// TIA Portal V20 export
// export: Created 2026-10-19T18:01:35.4601049Z, ExportSetting None, DisplayName Totally Integrated Automation Portal, DisplayVersion V20 Update 6, DisplayName TIA Portal Openness, DisplayVersion V20 Update 6, DisplayName TIA Portal Version Control Interface, DisplayVersion V20 Update 6, DisplayName SINAMICS Startdrive Advanced, DisplayVersion V20 SP1, DisplayName SINAMICS Startdrive G130, G150, S120, S150, SINAMICS MV, G220, S200, S210, DisplayVersion V20 SP1, DisplayName SINAMICS Startdrive G110M, G120, G120C, G120D, G120P, G115D, DisplayVersion V20 SP1, DisplayName STEP 7 Professional, DisplayVersion V20 Update 6, DisplayName STEP 7 Safety, DisplayVersion V20 Update 2, DisplayName WinCC Basic/Comfort/Advanced, DisplayVersion V20 Update 6, DisplayName WinCC Unified, DisplayVersion V20 Update 6
VAR_GLOBAL   // PLC tag table "Default tag table"
   Global_Estop AT %M1038.0 : Bool;
   Global_Estop_Error AT %M1038.1 : Bool;
   Mode_Change AT %IW502 : Int;
   Mode_Current AT %IW504 : Int;
   Reset_All AT %M510.2 : Bool;
   VTD_Buffers_In_Automatic AT %M510.1 : Bool;
   VTD_Automatic_Button AT %M510.0 : Bool;
   OPC_Enable AT %M11.6 : Bool;
   Mode_Change_2 AT %MW82 : UInt;
   MQTT_Enable AT %M11.7 : Bool;
   System_Byte AT %MB1 : Byte;
   FirstScan AT %M1.0 : Bool;
   DiagStatusUpdate AT %M1.1 : Bool;
   AlwaysTRUE AT %M1.2 : Bool;
   AlwaysFALSE AT %M1.3 : Bool;
   Clock_Byte AT %MB0 : Byte;
   Clock_10Hz AT %M0.0 : Bool;
   Clock_5Hz AT %M0.1 : Bool;
   "Clock_2.5Hz" AT %M0.2 : Bool;
   Clock_2Hz AT %M0.3 : Bool;
   "Clock_1.25Hz" AT %M0.4 : Bool;
   Clock_1Hz AT %M0.5 : Bool;
   "Clock_0.625Hz" AT %M0.6 : Bool;
   "Clock_0.5Hz" AT %M0.7 : Bool;
   Error_Word_1 AT %MW2001 : Word;
   Reintegration AT %M2000.3 : Bool;
   Charger_1st AT %Q106.1 : Bool;
   Charger_2nd AT %Q106.2 : Bool;
   Charger_3rd AT %Q106.3 : Bool;
   Reset_Comissioning AT %M2.0 : Bool;
   Tag_1 AT %IW384 : Int;
   Tag_2 AT %QW384 : Int;
   Carrousel_In_Automatic AT %M2.1 : Bool;
   Carrousel_Automatic_Button AT %M2.2 : Bool;
   State_PS AT %MW42 : Int;
   Debug_Barcode AT %M5.4 : Bool;
   mm_per_pulse AT %M300.0 : LReal;
   AE_Offset AT %MD104 : DInt;
   AE_Process_Offset AT %MD108 : Real;
   Safe_Mode AT %M9.6 : Bool;
   Dbug AT %M9.4 : Bool;
   Auto_Start_Barcode AT %M9.7 : Bool;
   Auto_Stop_Barcode AT %M9.5 : Bool;
END_VAR
VAR_GLOBAL CONSTANT   // user constants
   "Gross weight – rounded" : Byte := 0;   // Gross weight – rounded
   "Gross weight – rounded(1)" : Byte := 1;   // Gross weight – rounded
   "Tare weight – rounded" : Byte := 2;   // Tare weight – rounded
   "Net weight – rounded" : Byte := 3;   // Net weight – rounded
   "Gross weight – internal resolution" : Byte := 5;   // Gross weight – internal resolution
   "Tare weight – internal resolution" : Byte := 6;   // Tare weight – internal resolution
   "Net weight – internal resolution" : Byte := 7;   // Net weight – internal resolution
   Rate : Byte := 8;   // Rate – change in gross weight over time (in internal)
   "Weight unit" : Byte := 9;   // Weight unit (number representing unit from chart)
   Constant_1 : Int := 16;   // Gross weight of each POWERCELL in displayed
   Constant_2 : Int := 17;   // Net weight of each POWERCELL in displayed
   Constant_3 : Int := 18;   // Set threshold for customer overload xx d
   Constant_4 : Int := 218;   // Set threshold for customer overload xx d
   Constant_5 : Int := 19;   // Set threshold for customer underload xx D
   Constant_6 : Int := 219;   // Set threshold for customer underload xx D
   Constant_7 : Int := 40;   // Report/Write comparator 1 limit
   Constant_8 : Int := 240;   // Report/Write comparator 1 limit
   Constant_9 : Int := 41;   // Report / Write Comparator 1 High Limit
   Constant_10 : Int := 241;   // Report / Write Comparator 1 High Limit
   Constant_11 : Int := 42;   // Report/Write comparator 2 limit
   Constant_12 : Int := 242;   // Report/Write comparator 2 limit
   Constant_13 : Int := 43;   // Report / Write Comparator 2 High Limit
   Constant_14 : Int := 243;   // Report / Write Comparator 2 High Limit
   Constant_15 : Int := 44;   // Report/Write comparator 3 limit
   Constant_16 : Int := 244;   // Report/Write comparator 3 limit
   Constant_17 : Int := 45;   // Report / Write Comparator 3 High Limit
   Constant_18 : Int := 245;   // Report / Write Comparator 3 High Limit
   Constant_19 : Int := 46;   // Report/Write comparator 4 limit
   Constant_20 : Int := 246;   // Report/Write comparator 4 limit
   Constant_21 : Int := 47;   // Report / Write Comparator 4 High Limit
   Constant_22 : Int := 247;   // Report / Write Comparator 4 High Limit
   Constant_23 : Int := 48;   // Report/Write comparator 5 limit
   Constant_24 : Int := 248;   // Report/Write comparator 5 limit
   Constant_25 : Int := 49;   // Report / Write Comparator 5 High Limit
   Constant_26 : Int := 249;   // Report / Write Comparator 5 High Limit
   Constant_27 : Int := 50;   // Report/Write comparator 6 limit
   Constant_28 : Int := 250;   // Report/Write comparator 6 limit
   Constant_29 : Int := 51;   // Report / Write Comparator 6 High Limit
   Constant_30 : Int := 251;   // Report / Write Comparator 6 High Limit
   Constant_31 : Int := 52;   // Report/Write comparator 7 limit
   Constant_32 : Int := 252;   // Report/Write comparator 7 limit
   Constant_33 : Int := 53;   // Report / Write Comparator 7 High Limit
   Constant_34 : Int := 253;   // Report / Write Comparator 7 High Limit
   Constant_35 : Int := 54;   // Report/Write comparator 8 limit
   Constant_36 : Int := 254;   // Report/Write comparator 8 limit
   Constant_37 : Int := 55;   // Report / Write Comparator 8 High Limit
   Constant_38 : Int := 255;   // Report / Write Comparator 8 High Limit
   Constant_39 : Int := 95;   // Report/Write Zero adjustment count
   Constant_40 : Int := 295;   // Report/Write Zero adjustment count
   Constant_41 : Int := 201;   // Write Preset tare (display unit) Parameter: Pre–tare weight (float 32) placed in Measuring value
   Constant_42 : Int := 400;   // Tare when stable
   Constant_43 : Int := 401;   // Zero when stable
   Constant_44 : Int := 402;   // Clear tare
   Constant_45 : Int := 403;   // Tare immediately
   Constant_46 : Int := 404;   // Zero immediately
   Constant_47 : Int := 410;   // Trigger ePrint (Trigger Alibi Memory)
   Constant_48 : Int := 510;   // Apply Comparators
   Constant_49 : Int := 1000;   // Force all outputs OFF
   Constant_50 : Int := 1900;   // Alarm bit – write value of bit when in test mode
   Constant_51 : Int := 1901;   // Motion bit – write value of bit when in test mode
   Constant_52 : Int := 1902;   // Net mode bit – write value of bit when in test mode
   Constant_53 : Int := 1903;   // Center of zero bit – write value of bit when in test mode
   Constant_54 : Int := 1904;   // Alt weight bit – write value of bit when in test mode
   Constant_55 : Int := 1905;   // Device bit 1 – write value of bit when in test mode
   Constant_56 : Int := 1906;   // Device bit 2– write value of bit when in test mode
   Constant_57 : Int := 1907;   // Device bit 3– write value of bit when in test mode
   Constant_58 : Int := 1908;   // Device bit 4– write value of bit when in test mode
   Constant_59 : Int := 1909;   // Device bit 5– write value of bit when in test mode
   Constant_60 : Int := 1910;   // Device bit 6– write value of bit when in test mode
   Constant_61 : Int := 1911;   // Device bit 7– write value of bit when in test mode
   Constant_62 : Int := 1912;   // Performance Mode Parameter: 0 – send performance count at A/D rate 1 – send performance count at 1 ms interval n – send performance count at n ms interval
   Constant_63 : Int := 2000;   // No operation command – used to test command
   Constant_64 : Int := 2002;   // Continue to next step in sequence
   Constant_65 : Int := 2003;   // Continue to next step in sequence
   Constant_66 : Int := 2004;   // Abort sequence … response value means abort in process
   Constant_67 : Int := 2005;   // After step failure, retries previous step in sequence
   Constant_68 : Int := 2006;   // After step failure, skips step and advances to next in sequence
   Constant_69 : Int := 2045;   // Step successful, next value
   Constant_70 : Int := 2046;   // Step successful
   Constant_71 : Int := 2047;   // Command has been received and is being evaluated (in process)
END_VAR
